Fanuc KAREL source: KT00323.KL

PROGRAM KT00323
%NOLOCKGROUP
VAR
  P1: JOINTPOS
  P2: POSITION
  OUT: BOOLEAN
BEGIN
  OUT = P1 <> P2
END KT00323
